TYPE "ST_SequenceStep"
VERSION : 0.1
   STRUCT
      Visited : Bool;
      LastDuration : Time;
      ErrorActive : Bool;
      WarningActive : Bool;
   END_STRUCT;

END_TYPE

